DATA_BLOCK "db160_BC400_SetupPorTensao"
TITLE = db160_BC400_SetupPorTensao (DB160)
{ S7_Optimized_Access := 'FALSE' }
AUTHOR : 'Reginaldo Lobo'
VERSION : 0.2
////====================================
//// db160_BC400_SetupPorTensao (DB160)
//// O QUE FAZ : guarda os valores SALVOS do Setup de cada chave do banco BC400 (13 chaves, ate 16 posicoes),
////             SEPARADOS POR CHAVEAMENTO do banco (1 = 220 V, 2 = 380 V, 3 = 440 V). Cada linha de
////             tabela e um chaveamento; cada coluna e uma chave.
//// POR QUE EXISTE : a resistencia das chaves e a mesma nas 3 tensoes (informado pelo usuario em 25/10/2026),
////             logo o kW real de cada chave MUDA com a tensao (P = V^2 / R). O DB158 (setup.kwReal[]) guarda um
////             unico valor por chave, sem dizer em que tensao foi medido. Este DB guarda um valor por chave
////             E por tensao, mais a tensao e a base (kW sem carga) usadas no instante do Salvar.
//// ESCRITOR  : FB100 v0.3 (fb100_setupChaves) na borda de subida de ComandoSalvar, na linha do chaveamento
////             ativo (selV.tensaoSel). O chaveamento ativo e INFORMADO PELO HTML/Node-RED (decisao do usuario em
////             25/10/2026: "Pelo HTML/Node-red") - o PLC nao mede nem deduz. Leitor: Node-RED/HTML (v2.5 / v1.9.78).
//// POR QUE DB GLOBAL SEM OTIMIZACAO : leitura por offset fixo via S7 (PUT/GET) pelo Node-RED, igual ao DB158.
//// NAO TOCA no DB158: nenhum offset do DB158 muda; o Node-RED v2.4 continua valendo.
//// NUMERACAO : DB160 = base do banco (158) + 2 = "reserva +2" do gabarito de banco em
////             claude/PLANO_NUMERACAO_BLOCOS_PLC.md. NAO conflita com DB163 (instancia FB101). Registrar na
////             aba "Blocos_novos" da planilha PLANO_NUMERACAO_BLOCOS_PLC.
//// INDICES   : primeiro indice = chaveamento (1 = 220 V, 2 = 380 V, 3 = 440 V); segundo indice = chave (1..16).
////             Posicao linear p = (chaveamento - 1) * 16 + (chave - 1)   (0..47)
//// OFFSETS (ASSUMIDOS, conferir na coluna "Deslocamento" do TIA apos compilar - nao foi compilado):
////    setupV.tensaoV[1..3]        DBW0, DBW2, DBW4                (constantes 220, 380, 440)
////    setupV.kwReal[c,k]          DBD6   + 4  * p   (Real, kW real = kW com a chave - base)
////    setupV.rMedidoOhm[c,k]      DBD198 + 4  * p   (Real, ohm equivalente em estrela por fase = V^2 / (kW real * 1000))
////    setupV.vMedidaV[c,k]        DBD390 + 4  * p   (Real, tensao media fase-fase no instante do Salvar)
////    setupV.baseKw[c,k]          DBD582 + 4  * p   (Real, kW sem carga usado no Salvar)
////    setupV.setupData[c,k]       DBB774 + 12 * p   (DTL, data/hora do Salvar)
////    setupV.setupOk[c,k]         DBX1350.0 + p     (Bool, byte 1350 + p/8, bit p mod 8)
////    selV.tensaoSel              DBW1356           (Int, NOVO v0.2: chaveamento ativo informado pelo HTML/Node-RED:
////                                                   0 = nao informado, 1 = 220 V, 2 = 380 V, 3 = 440 V)
//// ATENCAO RETENTIVIDADE : estes valores precisam sobreviver a reinicio da CPU. Conferir no TIA (propriedades do DB)
////             que o DB esta retentivo. O DB158 esta como NON_RETAIN - pergunta pendente, nao alterada aqui.
//// ATENCAO DOWNLOAD : DB nao otimizado novo = carga inicial sem perda de dados existentes (DB novo).
//// v0.1 (25/10/2026): criacao. Nao compilado no TIA. Nao testado em hardware.
//// v0.2 (25/10/2026): + selV.tensaoSel (chaveamento ativo, escrito pelo Node-RED rota /tensao). Membro novo no FIM:
////             nenhum offset da v0.1 mudou. Se a v0.1 JA foi baixada no PLC, baixar a v0.2 REINICIALIZA o DB (DB
////             nao otimizado com membro novo) - ainda sem valores de Setup nele, entao nada se perde.
//// NAO ha 'tensao de referencia' (V_ref) no DB: ela e desconhecida e sera descoberta na pratica pelo Setup
////             (decisao do usuario em 25/10/2026). Por isso o R teorico NAO e gravado aqui.
//// Fonte: claude/ESPECIFICACAO_CARD_CHAVES_DB55_FB200.md (secao 4 e 7) + claude/PLANO_NUMERACAO_BLOCOS_PLC.md
////=====================================
   VAR
      setupV : Struct
         tensaoV     : Array[1..3] of Int;              // identificacao de cada chaveamento: 220, 380, 440 (V)
         kwReal      : Array[1..3, 1..16] of Real;      // kW real de cada chave naquele chaveamento
         rMedidoOhm  : Array[1..3, 1..16] of Real;      // ohm equivalente em estrela por fase (V^2 / (kW real * 1000))
         vMedidaV    : Array[1..3, 1..16] of Real;      // tensao media fase-fase no instante do Salvar (V)
         baseKw      : Array[1..3, 1..16] of Real;      // kW sem carga (BaseKW) usado no Salvar
         setupData   : Array[1..3, 1..16] of DTL;       // data/hora do Salvar (RD_SYS_T)
         setupOk     : Array[1..3, 1..16] of Bool;      // TRUE = esta chave tem Setup salvo neste chaveamento
      END_STRUCT;
      selV : Struct
         tensaoSel   : Int;                             // chaveamento ativo informado pelo HTML/Node-RED: 0 = nao informado, 1 = 220 V, 2 = 380 V, 3 = 440 V
      END_STRUCT;
   END_VAR


BEGIN
   setupV.tensaoV[1] := 220;
   setupV.tensaoV[2] := 380;
   setupV.tensaoV[3] := 440;
   selV.tensaoSel := 0;   // chaveamento NAO informado ate o operador escolher no HTML
   // demais membros: 0 / FALSE (sem Setup salvo). 14..16: reservado.

END_DATA_BLOCK
